// ============================================================================
// OB123.scl - TIA导入样例 主组织块 (全工站结构体整块传递架构)
// ============================================================================
// 描述:
//   DJ-2026-901 TIA导入样例 PLC 控制系统主循环调度程序.
//   全工站通过 VAR_IN_OUT 结构体整块传递 (Struct Chunk Passing), 遵循 LSP-905 规范.
//   每个功能块通过自己的背景 DB 单实例调用 (TIA 全局 DB 不能放 FB 实例, LSP-905 §4.11);
//   VAR_IN_OUT 按引用传递, 调用后不需要再把结构体写回 GlobalVars_DJ2026901.
//
// 块名与编号 (LSP-905 §3.4/§4.11):
//   块名带项目标记 DJ2026901, 不叫 Main/OB1, 导入时不会覆盖你项目里已有的同名块.
//   主程序固定 OB123; TIA 从源生成块时自己分配块号, 源文件里写不了 (TIA V19 实测), 导入后必须在 TIA 里手工改成 OB123 (见 程序架构文档 §7.4).
//   如果你的项目已有主程序, 也可以不导入本 OB, 只把下面几行调用复制进你自己的主程序.
//   每个工位一行调用, 工位清单在建项目时由 project create --station 给出 (CHG-SCPT-2026-635).
// ============================================================================
ORGANIZATION_BLOCK "DJ2026901_Main"
{ S7_Optimized_Block := 'TRUE' }
VERSION : 1.0

VAR_TEMP
END_VAR

BEGIN
    // ============================================================================
    // 第1部分：外部设备交互 (ST_3001_ExternalDevice)
    // ============================================================================
    "DB_3001_ExternalInteraction_DJ2026901"(io_stExternal := "GlobalVars_DJ2026901".stExternal);

    // ============================================================================
    // 第2部分：工位动作机构 (ST_1001_Station1), 每个工位一个背景 DB
    // ============================================================================
    "DB_1001_Station1_DJ2026901"(io_stStation := "GlobalVars_DJ2026901".stStation1);
    "DB_1001_Station2_DJ2026901"(io_stStation := "GlobalVars_DJ2026901".stStation2);
    "DB_1001_Station3_DJ2026901"(io_stStation := "GlobalVars_DJ2026901".stStation3);

    // ============================================================================
    // 第3部分：公共报警与 OMAC 状态机 (ST_2001_CommonAlarm)
    // ============================================================================
    "DB_2001_CommonAlarm_DJ2026901"(io_stGlobal := "GlobalVars_DJ2026901".stGlobal);

END_ORGANIZATION_BLOCK
